// I_Axis - what the RBG sequence needs from a positioning axis, whatever
// drives it: the simulated FB_Axis or the NC axis FB_AxisNc. Units are metres.
INTERFACE I_Axis

// Drive to an absolute position: eBusy while moving, eDone in position, eError on a fault.
METHOD MoveAbs : E_CmdResult
VAR_INPUT
    lrPos : LREAL;   // target [m]
END_VAR
END_METHOD

// Acknowledge a fault: the axis stops where it is and waits for a new target.
METHOD Reset
VAR_INPUT
END_VAR
END_METHOD

// Stop now (end of a jog, stop mode). The axis then waits for a new target.
METHOD Halt
VAR_INPUT
END_VAR
END_METHOD

// Actual position [m].
PROPERTY ActPos : LREAL
GET
END_GET
END_PROPERTY

PROPERTY Error : BOOL
GET
END_GET
END_PROPERTY

END_INTERFACE

(* stored: Version 1.1.0.1
   Itf I_Axis: Id {9b28e949-89ed-5419-a7f0-9a6bdce1367e}
   Method MoveAbs: Id {dd794198-a322-f627-73c3-ee0aa6a0c16f}
   Method Reset: Id {d3d6b18d-834b-8472-c693-07475f06f462}
   Method Halt: Id {b74cdb8b-123b-8062-9273-8f6dca2dddd3}
   Property ActPos: Id {b3a11f7d-a42f-8622-f90c-767f67eecf59}
   Get Get: Id {73ab3f9e-b2ff-23b8-ea5a-12563a4a9198}
   Property Error: Id {1f9964c6-7b7f-7b69-ab3a-ac49e291e8e6}
   Get Get: Id {7cc6907c-8455-c086-fdb3-a496d367986f} *)
